FUNCTION_BLOCK CompositeTest (* Composite FB containing a basic FB *)
  (* Standard: 61499-1; Description: Copyright (c) 2026 Martin Erich Jobst This program and the accompanying materials are made available under the terms of the Eclipse Public License 2.0 which is available at https://www.eclipse.org/legal/epl-2.0/ SPDX-License-Identifier: EPL-2.0 *)
  (* Version 1.0, 2026-10-23, Martin Jobst *)
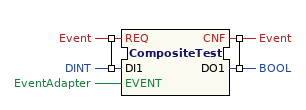
  EVENT_INPUT
    REQ WITH DI1; (* Request *)
  END_EVENT
  EVENT_OUTPUT
    CNF WITH DO1; (* Confirmation *)
  END_EVENT
  VAR_INPUT
    DI1 : DINT := DINT#42;
  END_VAR
  VAR_OUTPUT
    DO1 : BOOL;
  END_VAR
  SOCKETS
    EVENT : EventAdapter; (* Event/data adapter *)
  END_SOCKETS
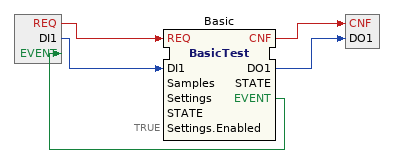
  (* Group ControlGroup: Grouped example *) {SET_ATTRIBUTE(IntegerAttribute, 2)}
  (* Composite network comment *)
  FBS
    Basic : fixture::basic::BasicTest(Settings.Enabled := TRUE {SET_ATTRIBUTE(IntegerAttribute, 3)}); {SET_ATTRIBUTE(GroupName, ControlGroup)}
  END_FBS
  EVENT_CONNECTIONS
    REQ TO Basic.REQ; (* Request forwarding *)
    Basic.CNF TO CNF;
  END_CONNECTIONS
  DATA_CONNECTIONS
    DI1 TO Basic.DI1;
    Basic.DO1 TO DO1;
  END_CONNECTIONS
  ADAPTER_CONNECTIONS
    Basic.EVENT TO EVENT;
  END_CONNECTIONS
END_FUNCTION_BLOCK
